FUNCTION_BLOCK tonrblock
VAR_INPUT
	in:BOOL;
	reset:BOOL;
	pt:TIME;
	
END_VAR
VAR_OUTPUT
	out:BOOL;
	et:TIME;
END_VAR
VAR
	tstarttime:TIME;
	tsavedtime:TIME;
	brunning:BOOL;
	
END_VAR

IF reset THEN
	tsavedtime:=T#0MS;
	et:=T#0MS;
	out:=FALSE;
	brunning:=FALSE;
ELSIF in THEN
     IF NOT brunning THEN
        tstarttime:=TIME();
        brunning:=TRUE;		 
	 END_IF
	 et:=tsavedtime+(TIME()-tstarttime);
	 IF et >= pt THEN;
		 et:=pt;
		 out:=TRUE;
	 END_IF
ELSE
	IF brunning THEN
		tsavedtime:=et;
		brunning:=FALSE;
	END_IF
END_IF

END_FUNCTION_BLOCK

(* stored: Version 1.1.0.1, ProductVersion 3.1.4024.16
   POU tonrblock: Id {04b5c1fe-71e6-4d87-80db-7edc957602dc}, SpecialFunc None *)
